Fanuc KAREL source: KT00941.KL

PROGRAM KT00941
%NOLOCKGROUP
VAR
  ENTRY: INTEGER
  PNAME: STRING[80]
  VNAME: STRING[80]
  STATUS: INTEGER
  VALUE: XYZWPREXT
BEGIN
  ENTRY = 0
  PNAME = ''
  VNAME = 'VALUE'
  GET_VAR(ENTRY, PNAME, VNAME, VALUE, STATUS)
END KT00941
